(* IEC 61131-3 sources: plc-st-test/packages/cli/test/fixtures/beckhoff-pointers/src, 2 files *)

(* ---- ST_Pair.st ---- *)
TYPE ST_Pair :
STRUCT
  nA : INT;
  nB : DINT;
END_STRUCT;
END_TYPE

(* ---- FB_Counter.st ---- *)
FUNCTION_BLOCK FB_Counter
VAR_OUTPUT
  nCount : INT;
END_VAR
METHOD Bump
  nCount := nCount + 1;
END_METHOD
END_FUNCTION_BLOCK
